// TIA Portal V20 export
FUNCTION_BLOCK "Drehtelleransteuerung"   // FB117, STL
TITLE = Drehteller Ansteuerung über Schütz, Abfrage Endschalter
{ S7_Optimized_Access := 'TRUE' }
// stored: AutoNumber false, MemoryReserve 100
   VAR_INPUT
      ES_GS : Bool;
      ES_Motor_aus : Bool;
      Automatik : Bool;
      Manuell : Bool;
      Einrichten : Bool;
      Ablauf_aktiv : Bool;
      Richten : Bool;
      SM_reset : Bool;
      Reset_Frg : Bool;
      Not_Aus_OK : Bool;
      Tueren_OK : Bool;
      Lichtvorhang_OK : Bool;
      Sicherheitsbit_DT : Bool;
      TP_Taste_tippen : Bool;
      Start_taste_tippen : Bool;
      links0_rechts1_drehen : Bool;
      Richten_erforderlich : Bool;
      LVZ_Timer : Timer;
      Timer_ueberdrehen : Timer;
      SVZ : Timer;
   END_VAR
   VAR_OUTPUT
      Schuetz_links : Bool;
      Schuetz_rechts : Bool;
      DT_Bremse : Bool;
   END_VAR
   VAR_IN_OUT
      Freigabe_DT : Bool;
      Manuellfreigabe : Bool;
      Richtenfreigabe : Bool;
      Fertigmeldung_Drehteller : Bool;
      Betriebsfertigmeldung : Bool;
      SM_GS : Bool;
      SM_AS : Bool;
      SM_Wartung : Bool;
      Auto_Frg_GS : Bool;
      Auto_Frg_AS : Bool;
      Manu_Frg_GS : Bool;
      Manu_Frg_AS : Bool;
      Einr_Frg_GS : Bool;
      Einr_Frg_AS : Bool;
      Init_Frg_GS : Bool;
      Init_Frg_AS : Bool;
      Richt_Frg_GS : Bool;
      Richt_Frg_AS : Bool;
   END_VAR
   VAR
      SchrittA1 : Bool;
      SchrittA2 : Bool;
      SchrittA3 : Bool;
      HM_DT_Frg_loeschen : Bool;
      FP_DT_frg_loeschen : Bool;
      SchrittM1 : Bool;
      SchrittM2 : Bool;
      LV_unterbrochen : Bool;
      HM_Tippen : Bool;
      FP_Tippen : Bool;
      FP_Start_Tippen : Bool;
   END_VAR
BEGIN

NETWORK
TITLE = Störmeldungen
      A     #ES_GS;
      A     #SchrittA1;
      AN    #SchrittA2;
      O(;
      AN    #ES_GS;
      A     #SchrittA2;
      AN    #SchrittA3;
      );
      AN    #SM_reset;
      L     S5T#1S;
      SD    #LVZ_Timer;

      A     #LVZ_Timer;
      S     #SM_GS;


      AN    #ES_Motor_aus;
      A     #SchrittA1;
      AN    #SchrittA2;
      O(;
      A     #ES_Motor_aus;
      A     #SchrittA2;
      AN    #SchrittA3;
      );
      O(;
      AN    #ES_GS;
      A     #ES_Motor_aus;
      );
      AN    #SM_reset;
      L     S5T#1S;
      SD    #Timer_ueberdrehen;

      A     #Timer_ueberdrehen;
      S     #SM_AS;

      A     #SM_GS;
      A     #SM_reset;
      R     #SM_GS;

      A     #SM_AS;
      A     #SM_reset;
      R     #SM_AS;



NETWORK
TITLE = Lichtvorhang unterbrochen speichern
      A     #SchrittA1;
      AN    #Lichtvorhang_OK;
      S     #LV_unterbrochen;
      R     #SchrittA1;
      R     #SchrittA1;
      R     #SchrittA3;
      R     #DT_Bremse;
      R     #Schuetz_rechts;
      R     #Schuetz_links;



NETWORK
TITLE = Fertigmeldung DT
      A     #Betriebsfertigmeldung;
      FP    #HM_DT_Frg_loeschen;
      =     #FP_DT_frg_loeschen;

      A     #FP_DT_frg_loeschen;
      S     #Fertigmeldung_Drehteller;
      R     #Betriebsfertigmeldung;



NETWORK
TITLE = Sicherheitsabfragen
      A     #Not_Aus_OK;
      A     #Tueren_OK;
      A     #Lichtvorhang_OK;
      A     #Sicherheitsbit_DT;
      JCN   Ende;
      A     #Automatik;
      A     #Ablauf_aktiv;
      O;
      A     #Manuell;
      A     #Manuellfreigabe;
      O     #Richten_erforderlich;
      JC    M010;
      A     #Manuell;
      AN    #Manuellfreigabe;
      JC    M050;

      JU    Ende;



NETWORK
TITLE = Schritt1: Ansteuerung DT Automatik/Manuell
M010: A     #SchrittA1;
      JC    M020;
      A     #Freigabe_DT;
      A     #ES_GS;
//   UN    #ES_Motor_aus
      O     #Manuellfreigabe;
      O(;
      A     #Richten_erforderlich;
      A     #Richtenfreigabe;
      );
      O(;
      A     #Lichtvorhang_OK;
      A     #LV_unterbrochen;
      );
      AN    #SM_GS;
      AN    #SM_AS;
      S     #DT_Bremse;
      R     #Freigabe_DT;
      R     #Richtenfreigabe;
      R     #LV_unterbrochen;

      A     #DT_Bremse;
      A     #links0_rechts1_drehen;
      S     #Schuetz_rechts;

      A     #DT_Bremse;
      AN    #links0_rechts1_drehen;
      S     #Schuetz_links;

      A     #Schuetz_rechts;
      O     #Schuetz_links;
      A     #DT_Bremse;
      S     #SchrittA1;
      JC    M021;
      BEU;
M021: CLR;
      SD    #SVZ;
      BEU;



NETWORK
TITLE = Schritt2: ES_GS geht weg
M020: A     #SchrittA2;
      JC    M030;
      AN    #ES_GS;
      A     #ES_Motor_aus;
      O     #SM_GS;
      O     #SM_AS;
      S     #SchrittA2;
      JC    M031;
      BEU;
M031: CLR;
      SD    #SVZ;
      BEU;



NETWORK
TITLE = Schritt3: ES_GS kommt und ES_Motor_aus geht weg
M030: A     #SchrittA3;
      JC    M040;
      A     #ES_GS;
      A     #ES_Motor_aus;
      AN    #Richten_erforderlich;
      O(;
      A     #ES_Motor_aus;
      A     #ES_GS;
      A     #Richten_erforderlich;
      );
      O     #SM_GS;
      O     #SM_AS;
      O(;
      AN    #SM_GS;
      AN    #SM_AS;
      A     #ES_GS;
      AN    #ES_Motor_aus;
      A     #SM_reset;
      );
      R     #Schuetz_rechts;
      R     #Schuetz_links;
      R     #DT_Bremse;
      S     #Betriebsfertigmeldung;
      S     #SchrittA3;
      JC    M041;
      BEU;
M041: CLR;
      SD    #SVZ;
      BEU;



NETWORK
TITLE = Schrittkettenende
M040: SET;
      R     #SchrittA1;
      R     #SchrittA2;
      R     #SchrittA3;
      R     #Manuellfreigabe;
      BEU;



NETWORK
TITLE = Schritt1: Ansteuerung DT Manuell-Tippen
M050: A     #TP_Taste_tippen;
      A     #Start_taste_tippen;
      FP    #FP_Start_Tippen;
      S     #HM_Tippen;

      A(;
      A     #ES_GS;
      A     #ES_Motor_aus;
      FP    #FP_Tippen;
      );
      ON    #TP_Taste_tippen;
      ON    #Start_taste_tippen;
      R     #HM_Tippen;

      A     #HM_Tippen;
      =     #DT_Bremse;

      A     #DT_Bremse;
      A     #links0_rechts1_drehen;
      =     #Schuetz_rechts;

      A     #DT_Bremse;
      AN    #links0_rechts1_drehen;
      =     #Schuetz_links;

      BEU;



NETWORK
TITLE = Ende wenn nichts angewählt
Ende: NOP   0;
      SET;
      R     #DT_Bremse;
      R     #Schuetz_rechts;
      R     #Schuetz_links;
      R     #SchrittA1;
      R     #SchrittA2;
      R     #SchrittA3;
      R     #Manuellfreigabe;

      BEU;

END_FUNCTION_BLOCK
